PROGRAM MAIN
VAR
    motorCtrlWord AT%Q* : UINT; // Motor ControlWord output
    loadCtrlWord AT%Q* : UINT; // Load ControlWord output
    motorStatWord AT%I* : UINT; // Motor StatusWord input
    loadStatWord AT%I* : UINT; // Load StatusWord input
    seqPlaybackDone AT%I* : BOOL; // Sequencer playback done (latched)
    experimentActiveOut AT%Q* : BOOL; // ModeManager experiment active output
    preArmOut AT%Q* : BOOL; // ModeManager logger pre-arm output
    resetOut AT%Q* : BOOL; // One-shot reset pulse output
    enableCurrentOut AT%Q* : BOOL; // Current enable gate output

    // FSM state
    modeState : E_ModeState := E_ModeState.IDLE;
    modeOutputs : ST_ModeOutputs;

    // Decoded request flags (from GVL_MODE.modeFlags)
    servoEnableReq : BOOL := FALSE;
    experimentStartReq : BOOL := FALSE;
    fbModeManagerCore : FB_ModeManagerCore;

    // Drive state
    driveReady : BOOL := FALSE;
    motorDriveReady : BOOL := FALSE;
    loadDriveReady : BOOL := FALSE;
    enableEffective : BOOL := FALSE;

    fbMotorStateMachine : FB_StateMachineControl;
    fbLoadStateMachine : FB_StateMachineControl;
    loggerReadyIn AT%I* : BOOL; // ExperimentLogger file FSM ACTIVE
    loggerFileReleasedIn AT%I* : BOOL; // ExperimentLogger close completed
    loggerErrorCodeIn AT%I* : UDINT; // ExperimentLogger session error
END_VAR

(* ===== 1. Decode input flags ===== *)
servoEnableReq := (GVL_MODE.modeFlags AND GVL_MODE.MODEF_SERVO_ENABLE) <> 0;
experimentStartReq := (GVL_MODE.modeFlags AND GVL_MODE.MODEF_EXPERIMENT_START_REQ) <> 0;

(* ===== 2. Request/watchdog/FSM core ===== *)
fbModeManagerCore(
    servoEnableRequest := servoEnableReq,
    experimentStartRequest := experimentStartReq,
    anyModeRequest := (GVL_MODE.modeFlags <> 0),
    resetRequest := GVL_MODE.resetReq,
    experimentActivePreviousScan := GVL_MODE.experimentActive,
    hostHeartbeatCounter := GVL_MODE.hostHeartbeatCounter,
    heartbeatTimeoutTicks := GVL_MODE.HEARTBEAT_TIMEOUT_TICKS,
    driveReadyPreviousScan := driveReady,
    loggerReady := loggerReadyIn,
    seqPlaybackDone := seqPlaybackDone
);

IF fbModeManagerCore.actions.consumeResetReq THEN
    GVL_MODE.resetReq := FALSE;
END_IF
IF fbModeManagerCore.actions.clearModeFlags THEN
    GVL_MODE.modeFlags := 0;
END_IF
IF fbModeManagerCore.actions.incrementResetAckCounter THEN
    GVL_MODE.resetAckCounter := GVL_MODE.resetAckCounter + 1;
END_IF
IF fbModeManagerCore.actions.incrementWatchdogTripCounter THEN
    GVL_MODE.watchdogTripCounter := GVL_MODE.watchdogTripCounter + 1;
END_IF

modeState := fbModeManagerCore.modeState;
enableEffective := fbModeManagerCore.driveEnable;

(* ===== 3. Drive state update ===== *)
fbMotorStateMachine(
    statusWord := motorStatWord,
    enable := enableEffective
);
fbLoadStateMachine(
    statusWord := loadStatWord,
    enable := enableEffective
);

motorCtrlWord := fbMotorStateMachine.controlWord;
loadCtrlWord := fbLoadStateMachine.controlWord;
motorDriveReady := (fbMotorStateMachine.driveState = E_DriveState.OPERATION_ENABLED);
loadDriveReady := (fbLoadStateMachine.driveState = E_DriveState.OPERATION_ENABLED);
driveReady := motorDriveReady AND loadDriveReady;

(* ===== 4. State-dependent outputs ===== *)
modeOutputs := F_DeriveModeOutputs(modeState := modeState);
experimentActiveOut := modeOutputs.experimentActiveOut;
preArmOut := modeOutputs.preArmOut;
resetOut := modeOutputs.resetOut;
enableCurrentOut := modeOutputs.enableCurrentOut;

GVL_MODE.experimentActive := experimentActiveOut;
IF modeState = E_ModeState.SERVO_READY THEN
    GVL_MODE.loggerFileReleased := FALSE;
    GVL_MODE.loggerErrorCode := 0;
ELSE
    GVL_MODE.loggerFileReleased := loggerFileReleasedIn;
    GVL_MODE.loggerErrorCode := loggerErrorCodeIn;
END_IF;
GVL_MODE.modeState := modeState;

END_PROGRAM

(* stored: Version 1.1.0.1
   POU MAIN: Id {9328c0c8-0c23-447b-8f8c-ef2a688ee9a0}, SpecialFunc None *)
